INTERFACE I_Meter EXTENDS I_Module

METHOD M_Cycle
END_METHOD

PROPERTY MeterState : ST_MeterState
GET
END_GET
END_PROPERTY

END_INTERFACE

(* stored: Version 1.1.0.1, ProductVersion 3.1.4024.15
   Itf I_Meter: Id {9db91630-56a0-4318-8827-292990481b53}
   Method M_Cycle: Id {03c77236-44e6-4291-97c3-44eeda3cafa6}
   Property MeterState: Id {082455e6-f72c-4a1f-8b92-f21d4ad7afa3}
   Get Get: Id {5844bdbe-7fb4-40b2-9186-60f735e69965} *)
